(* IEC 61131-3 sources: Lasal-MCP/examples/SampleSource/5_ClassInputOutputSolution/Stations/MachineControl/MachineControl/Class/_CheckOnlineStatus, 1 file *)

(* ---- _CheckOnlineStatus.st ---- *)
(*!
<Class
	Name               = "_CheckOnlineStatus"
	Revision           = "1.2"
	RealtimeTask       = "false"
	CyclicTask         = "true"
	DefCyclictime      = "50 ms"
	BackgroundTask     = "false"
	Sigmatek           = "true"
	OSInterface        = "false"
	HighPriority       = "false"
	Automatic          = "false"
	UpdateMode         = "Prescan"
	SharedCommandTable = "true"
	Objectsize         = "(600,180)"
	Comment            = "class for checking/alarming the online status">
	<Channels>
		<Server Name="AlarmState" Visualized="true" Initialize="false" WriteProtected="false" Retentive="false" Comment="actual status of the communication alarm"/>
		<Server Name="Locked" Visualized="false" Initialize="false" WriteProtected="true" Retentive="false" Comment="0 ... communication never was online&#13;&#10;1 ... communication was online"/>
		<Server Name="RestTime" Visualized="false" Initialize="false" WriteProtected="true" Retentive="false" Comment="rest time until alarm will be generated [millisec] (output)"/>
		<Client Name="AlarmCommunication" Required="true" Internal="true"/>
		<Client Name="AlarmNo" Required="true" Internal="false" Comment="alarm number for PLC offline alarm (input)"/>
		<Client Name="DelayTime" Required="true" Internal="false" DefValue="20000" Comment="delay time for alarm generating [millisec] (input)"/>
		<Client Name="toTCPComm" Required="true" Internal="false" Comment="Object channel to TCPCommunication."/>
	</Channels>
	<Dependencies>
		<Files>
			<File Path=".\Class\_CheckOnlineStatus\_CheckOnlineStatus_de.pdf"/>
			<File Path=".\Class\_CheckOnlineStatus\_CheckOnlineStatus_en.pdf"/>
		</Files>
	</Dependencies>
	<RevDoku>
		<Owner Company="Sigmatek"/>
		<Dokumentation Revision="1.2" Date="2016-11-04" Author="KaiAnd" Company="Sigmatek" Description="building the locked flag: Wait for first online status AND communication after system start (not only online status)&#13;&#10;also an optional timeDelay is implemented for the alarm generating"/>
		<Dokumentation Revision="1.1" Date="2016-10-10" Author="HubChr" Company="Sigmatek" Description="Added documentation pdfs."/>
		<Dokumentation Revision="1.0" Date="2015-06-24" Company="Sigmatek" Description="Creation."/>
	</RevDoku>
	<Network Name="_CheckOnlineStatus">
		<!-- List of Components in this network -->
		<Components>
			<Object
				Name       = "AlarmCommunication"
				Class      = "_AlarmX0Para"
				Position   = "(210,240)"
				Visualized = "true">
				<Channels>
					<Server Name="ClassSvr"/>
					<Client Name="Acknow"/>
					<Client Name="Config" Value="0"/>
					<Client Name="Group"/>
				</Channels>
			</Object>
		</Components>
		<Comments>
		</Comments>
		<!-- List of Connections in this network -->
		<Connections>
			<Connection Source="AlarmCommunication.Config" Destination="this.AlarmNo" Vertices="(210,330),(38,270),"/>
			<Connection Source="this.AlarmState" Destination="AlarmCommunication.ClassSvr" Vertices="(682,270),(510,330),"/>
			<Connection Source="this.AlarmCommunication" Destination="AlarmCommunication.ClassSvr"/>
		</Connections>
		<!-- Headerfiles -->
		<Options>
		</Options>
	</Network>
</Class>
*)
_CheckOnlineStatus : CLASS
  //Servers:
	Locked 	: SvrChCmd_DINT;
	AlarmState 	: SvrCh_DINT;
	RestTime 	: SvrCh_UDINT;
  //Clients:
	toTCPComm 	: CltChCmd_TCPCommunication;
	AlarmNo 	: CltCh_DINT;
	AlarmCommunication 	: CltChCmd__AlarmX0Para;
	DelayTime 	: CltCh_UDINT;
  //Variables:
		TimeMarkAlarm 	: UDINT;
  //Functions:

	FUNCTION VIRTUAL GLOBAL CyWork
		VAR_INPUT
			EAX 	: UDINT;
		END_VAR
		VAR_OUTPUT
			state (EAX) 	: UDINT;
		END_VAR;

	FUNCTION VIRTUAL GLOBAL AlarmState::Read
		VAR_OUTPUT
			output (EAX) 	: DINT;
		END_VAR;

	FUNCTION VIRTUAL GLOBAL AlarmState::Write
		VAR_INPUT
			input (EAX) 	: DINT;
		END_VAR
		VAR_OUTPUT
			result (EAX) 	: DINT;
		END_VAR;
  //Tables:
	FUNCTION @STD
		VAR_OUTPUT
			ret_code	: CONFSTATES;
		END_VAR;
	FUNCTION GLOBAL TAB @CT_;
END_CLASS;

#pragma using _AlarmX0Para
#pragma usingLtd TCPCommunication

FUNCTION VIRTUAL GLOBAL _CheckOnlineStatus::CyWork
	VAR_INPUT
		EAX 	: UDINT;
	END_VAR
	VAR_OUTPUT
		state (EAX) 	: UDINT;
	END_VAR
  VAR
  	myOnlineWarning : DINT;
  	myOnlineAlarm   : DINT;
  END_VAR

  //-----------------------------------------------------------------
  //  INIT
  //-----------------------------------------------------------------
  DelayTime := DelayTime.Read();
  myOnlineWarning := 0;
  myOnlineAlarm   := 0;

  //-----------------------------------------------------------------
  //  Online-Alarm:
  //-----------------------------------------------------------------

  // online and communication ... Status OK!
  if ( (toTCPComm.Online <> 0) &
       (toTCPComm.TransferRateReceive <> 0) ) then
    Locked := 1;      // Communication was online after system start

//  elsif (locked = 1) then
  else
    myOnlineWarning := 1;
  end_if;

  //-----------------------------------------------------------------
  //  building the alarm with delayTimer
  //-----------------------------------------------------------------

  // no online warning
  if (myOnlineWarning = 0) then
    TimeMarkAlarm := ops.tAbsolute;

  // online warning!
  else
    // time delay
    if ((ops.tAbsolute - TimeMarkAlarm) >= DelayTime) then
      myOnlineAlarm := 1;   // set alarm
    end_if;
  end_if;

  // write status to alarm server
  if (AlarmCommunication.ClassSvr.Read() <> myOnlineAlarm) then
    AlarmCommunication.ClassSvr.Write(input:=myOnlineAlarm);
  end_if;

  // write rest time to server
  RestTime := DelayTime - (ops.tAbsolute - TimeMarkAlarm);
  if (RestTime$DINT < 0) then
    RestTime := 0;
  end_if;

  //-----------------------------------------------------------------

	state := READY;

END_FUNCTION

FUNCTION VIRTUAL GLOBAL _CheckOnlineStatus::AlarmState::Read
	VAR_OUTPUT
		output (EAX) 	: DINT;
	END_VAR

	AlarmState := AlarmCommunication.ClassSvr.Read();
	output := AlarmState;

END_FUNCTION

FUNCTION VIRTUAL GLOBAL _CheckOnlineStatus::AlarmState::Write
	VAR_INPUT
		input (EAX) 	: DINT;
	END_VAR
	VAR_OUTPUT
		result (EAX) 	: DINT;
	END_VAR

	AlarmState := input;
	result := (AlarmCommunication.ClassSvr.Write(AlarmState))$DINT;

END_FUNCTION
